SUBAPPLICATION Uebung_253_AX (* Section-Switcher QUARTER, 8 Sections je eine auf Q1-Q8, Start alle aus *)
  (* Standard: 61499-2; Description: Copyright (c) 2026 Meisterschulen am Ostbahnhof This program and the accompanying materials are made available under the terms of the Eclipse Public License 2.0 which is available at https://www.eclipse.org/legal/epl-2.0/ SPDX-License-Identifier: EPL-2.0 *)
  (* Version 1.0, 2026-11-05, Franz Höpfinger, Meisterschulen am Ostbahnhof, initial API and implementation and/or initial documentation *)
  PACKAGE Uebungen;
  IMPORT logiBUS::io::DI::logiBUS_DI::Input_I1;
  IMPORT logiBUS::io::DI::logiBUS_DI::Input_I2;
  IMPORT logiBUS::io::DI::logiBUS_DI::Input_I7;
  IMPORT logiBUS::io::DI::logiBUS_DI::Input_I8;
  IMPORT logiBUS::io::DI::logiBUS_DI_Events::BUTTON_SINGLE_CLICK;
  IMPORT logiBUS::io::DQ::logiBUS_DO::Output_Q1;
  IMPORT logiBUS::io::DQ::logiBUS_DO::Output_Q2;
  IMPORT logiBUS::io::DQ::logiBUS_DO::Output_Q3;
  IMPORT logiBUS::io::DQ::logiBUS_DO::Output_Q4;
  IMPORT logiBUS::io::DQ::logiBUS_DO::Output_Q5;
  IMPORT logiBUS::io::DQ::logiBUS_DO::Output_Q6;
  IMPORT logiBUS::io::DQ::logiBUS_DO::Output_Q7;
  IMPORT logiBUS::io::DQ::logiBUS_DO::Output_Q8;
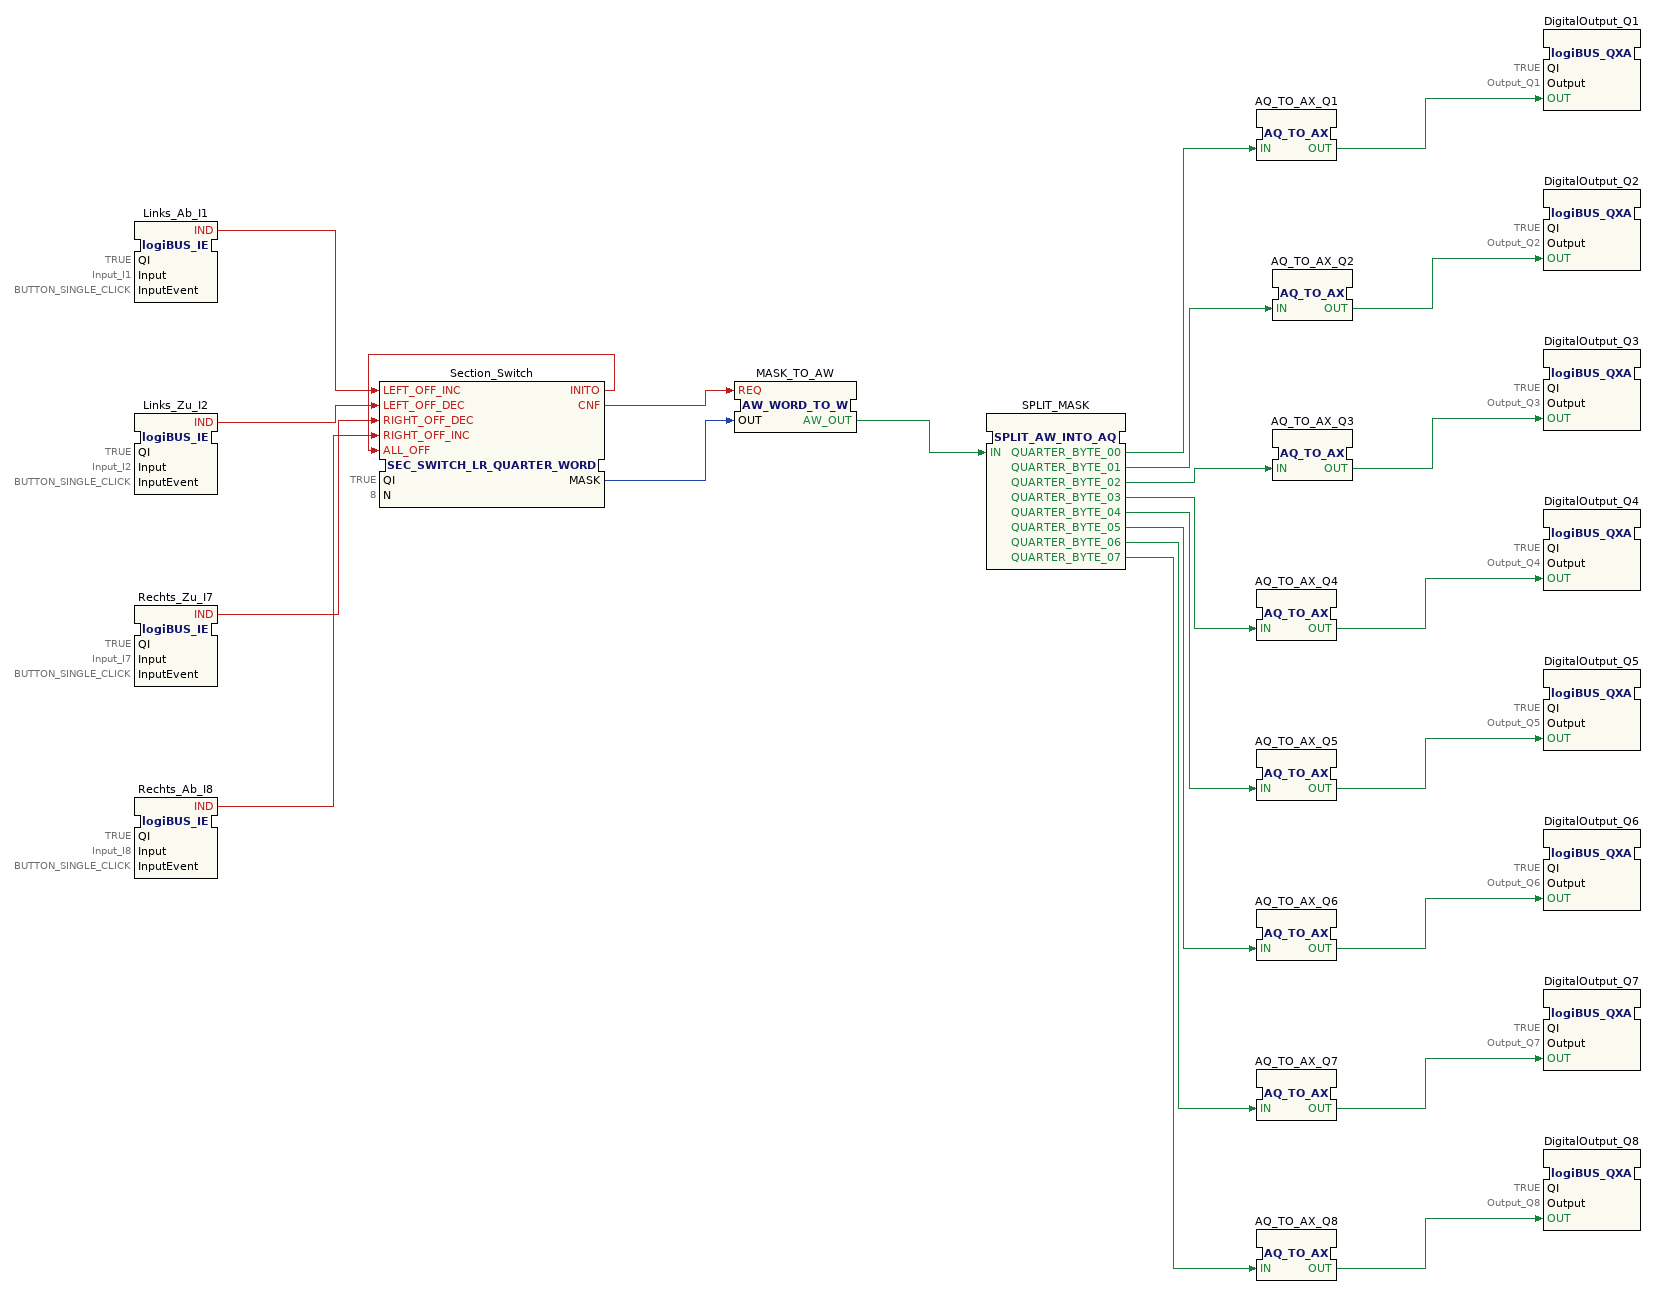
  FBS
    Links_Ab_I1 : logiBUS::io::DI::logiBUS_IE(QI := TRUE, Input := Input_I1, InputEvent := BUTTON_SINGLE_CLICK);
    Links_Zu_I2 : logiBUS::io::DI::logiBUS_IE(QI := TRUE, Input := Input_I2, InputEvent := BUTTON_SINGLE_CLICK);
    Rechts_Zu_I7 : logiBUS::io::DI::logiBUS_IE(QI := TRUE, Input := Input_I7, InputEvent := BUTTON_SINGLE_CLICK);
    Rechts_Ab_I8 : logiBUS::io::DI::logiBUS_IE(QI := TRUE, Input := Input_I8, InputEvent := BUTTON_SINGLE_CLICK);
    Section_Switch : logiBUS::sections::SEC_SWITCH_LR_QUARTER_WORD(QI := TRUE, N := 8); (* Startet sicher: INITO auf ALL_OFF, alle Sections aus *)
    MASK_TO_AW : adapter::conversion::unidirectional::AW_WORD_TO_W;
    SPLIT_MASK : adapter::splitting::SPLIT_AW_INTO_AQ;
    AQ_TO_AX_Q1 : adapter::conversion::unidirectional::AQ_TO_AX;
    DigitalOutput_Q1 : logiBUS::io::DQ::logiBUS_QXA(QI := TRUE, Output := Output_Q1);
    AQ_TO_AX_Q2 : adapter::conversion::unidirectional::AQ_TO_AX;
    DigitalOutput_Q2 : logiBUS::io::DQ::logiBUS_QXA(QI := TRUE, Output := Output_Q2);
    AQ_TO_AX_Q3 : adapter::conversion::unidirectional::AQ_TO_AX;
    DigitalOutput_Q3 : logiBUS::io::DQ::logiBUS_QXA(QI := TRUE, Output := Output_Q3);
    AQ_TO_AX_Q4 : adapter::conversion::unidirectional::AQ_TO_AX;
    DigitalOutput_Q4 : logiBUS::io::DQ::logiBUS_QXA(QI := TRUE, Output := Output_Q4);
    AQ_TO_AX_Q5 : adapter::conversion::unidirectional::AQ_TO_AX;
    DigitalOutput_Q5 : logiBUS::io::DQ::logiBUS_QXA(QI := TRUE, Output := Output_Q5);
    AQ_TO_AX_Q6 : adapter::conversion::unidirectional::AQ_TO_AX;
    DigitalOutput_Q6 : logiBUS::io::DQ::logiBUS_QXA(QI := TRUE, Output := Output_Q6);
    AQ_TO_AX_Q7 : adapter::conversion::unidirectional::AQ_TO_AX;
    DigitalOutput_Q7 : logiBUS::io::DQ::logiBUS_QXA(QI := TRUE, Output := Output_Q7);
    AQ_TO_AX_Q8 : adapter::conversion::unidirectional::AQ_TO_AX;
    DigitalOutput_Q8 : logiBUS::io::DQ::logiBUS_QXA(QI := TRUE, Output := Output_Q8);
  END_FBS
  EVENT_CONNECTIONS
    Links_Ab_I1.IND TO Section_Switch.LEFT_OFF_INC;
    Links_Zu_I2.IND TO Section_Switch.LEFT_OFF_DEC;
    Rechts_Zu_I7.IND TO Section_Switch.RIGHT_OFF_DEC;
    Rechts_Ab_I8.IND TO Section_Switch.RIGHT_OFF_INC;
    Section_Switch.INITO TO Section_Switch.ALL_OFF;
    Section_Switch.CNF TO MASK_TO_AW.REQ;
  END_CONNECTIONS
  DATA_CONNECTIONS
    Section_Switch.MASK TO MASK_TO_AW.OUT;
  END_CONNECTIONS
  ADAPTER_CONNECTIONS
    MASK_TO_AW.AW_OUT TO SPLIT_MASK.IN;
    SPLIT_MASK.QUARTER_BYTE_00 TO AQ_TO_AX_Q1.IN;
    AQ_TO_AX_Q1.OUT TO DigitalOutput_Q1.OUT;
    SPLIT_MASK.QUARTER_BYTE_01 TO AQ_TO_AX_Q2.IN;
    AQ_TO_AX_Q2.OUT TO DigitalOutput_Q2.OUT;
    SPLIT_MASK.QUARTER_BYTE_02 TO AQ_TO_AX_Q3.IN;
    AQ_TO_AX_Q3.OUT TO DigitalOutput_Q3.OUT;
    SPLIT_MASK.QUARTER_BYTE_03 TO AQ_TO_AX_Q4.IN;
    AQ_TO_AX_Q4.OUT TO DigitalOutput_Q4.OUT;
    SPLIT_MASK.QUARTER_BYTE_04 TO AQ_TO_AX_Q5.IN;
    AQ_TO_AX_Q5.OUT TO DigitalOutput_Q5.OUT;
    SPLIT_MASK.QUARTER_BYTE_05 TO AQ_TO_AX_Q6.IN;
    AQ_TO_AX_Q6.OUT TO DigitalOutput_Q6.OUT;
    SPLIT_MASK.QUARTER_BYTE_06 TO AQ_TO_AX_Q7.IN;
    AQ_TO_AX_Q7.OUT TO DigitalOutput_Q7.OUT;
    SPLIT_MASK.QUARTER_BYTE_07 TO AQ_TO_AX_Q8.IN;
    AQ_TO_AX_Q8.OUT TO DigitalOutput_Q8.OUT;
  END_CONNECTIONS
END_SUBAPPLICATION
